TYPE ST_PLCTONC :
STRUCT
	(* SDS *)
	stBaseDevice				:ST_BaseDeviceOut;

	(* SD6/SC6/SI6 *)
	stCIA402						:ST_CIA402Out;



(*



	dnReferencePosition			:DINT;			(* Value which is loaded as the actual position in the reference point. *)

*)
END_STRUCT
END_TYPE

(* stored: Version 1.1.0.1, ProductVersion 3.1.4024.15
   DUT ST_PLCTONC: Id {1920efb3-f853-4f9b-a4b4-a7fe07651d49} *)
